// SIMATIC S7-200 project (STEP 7-Micro/WIN), CPU 226 CN REL 02.01

SYMBOL_TABLE USUARIO1
act1             Q0.0
act2             Q0.1
act3             Q0.2
act4             Q0.3
act5             Q0.4
act6             Q0.5
act7             Q0.6
act8             Q0.7
act9             Q1.0
bot_verde        I2.5
bot_rojo         I2.4
selector         I2.7
QS               I2.6
END_SYMBOL_TABLE

ORGANIZATION_BLOCK PRINCIPAL:OB1
TITLE=COMENTARIOS DEL PROGRAMA
BEGIN
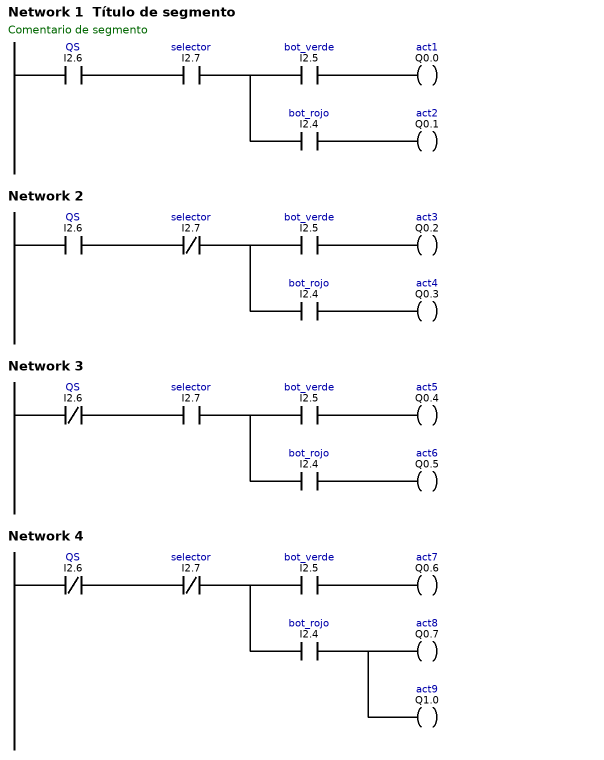
Network 1 // Título de segmento
// Comentario de segmento
LD     QS:I2.6
A      selector:I2.7
LPS
A      bot_verde:I2.5
=      act1:Q0.0
LPP
A      bot_rojo:I2.4
=      act2:Q0.1
Network 2
LD     QS:I2.6
AN     selector:I2.7
LPS
A      bot_verde:I2.5
=      act3:Q0.2
LPP
A      bot_rojo:I2.4
=      act4:Q0.3
Network 3
LDN    QS:I2.6
A      selector:I2.7
LPS
A      bot_verde:I2.5
=      act5:Q0.4
LPP
A      bot_rojo:I2.4
=      act6:Q0.5
Network 4
// (network saved uncompiled; LAD cells follow)
// row 0: c0 -|/|- QS:I2.6  c1 -|/|- selector:I2.7 v  c2 -| |- bot_verde:I2.5  c3 -( ) act7:Q0.6
// row 1: c1 ^  c2 -| |- bot_rojo:I2.4 v  c3 -( ) act8:Q0.7
// row 2: c2 ^  c3 -( ) act9:Q1.0
END_ORGANIZATION_BLOCK
